(* CODESYS project Controls.export

Project tree, tasks and I/O mapping:
  visualisation Controls
*)

// /Controls
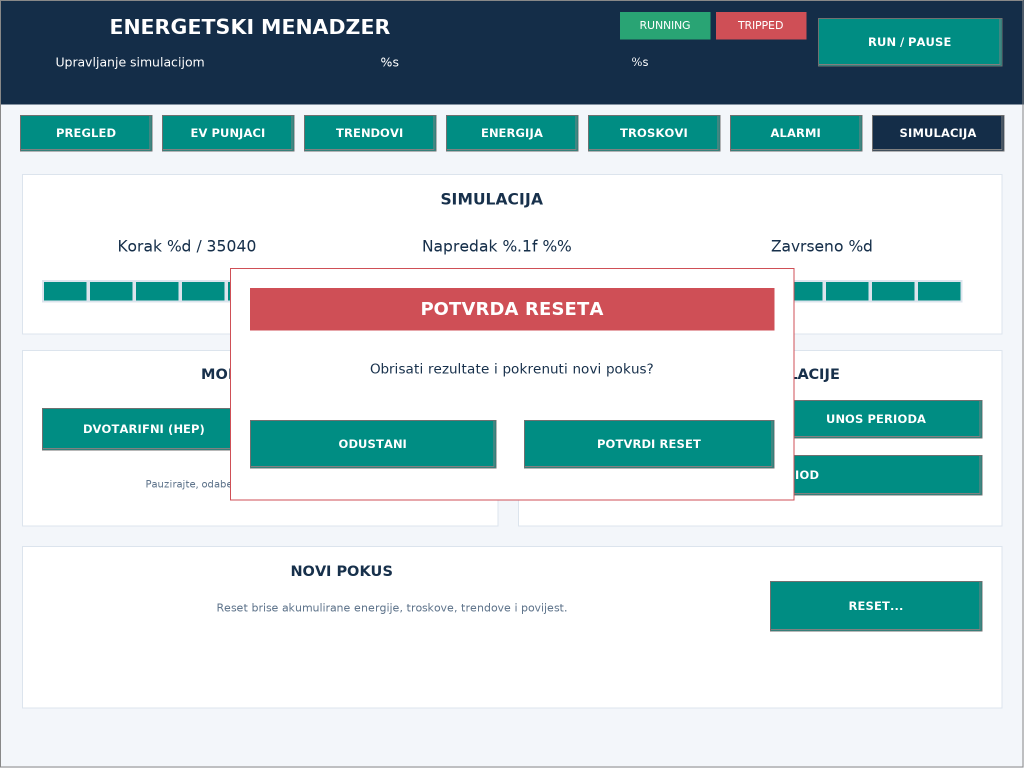
VISUALIZATION Controls  // 1024x768
    Rectangle (0,0 1024x768)
    Rectangle (0,0 1024x104)
    Rectangle (20,10 460x34), "ENERGETSKI MENADZER"
    Rectangle (20,48 220x28), "Upravljanje simulacijom"
    Rectangle (260,49 260x26), "%s", text variable: Team_HMI.sDateTime
    Rectangle (530,49 220x26), "%s", text variable: Team_HMI.sPriceMode
    Button (818,18 184x48), "RUN / PAUSE"
        toggle SimCtrl.run
    Rectangle (620,12 90x27), "PAUSED", invisible if: SimCtrl.run
    Rectangle (620,12 90x27), "RUNNING", invisible if: NOT SimCtrl.run
    Rectangle (716,12 90x27), "TRIPPED", invisible if: NOT SimCtrl.tripped
    Button (20,115 132x36), "PREGLED"
        OnMouseClick:  Assign=Overview, Type=Assignment
    Button (162,115 132x36), "EV PUNJACI"
        OnMouseClick:  Assign=EVs, Type=Assignment
    Button (304,115 132x36), "TRENDOVI"
        OnMouseClick:  Assign=Trends, Type=Assignment
    Button (446,115 132x36), "ENERGIJA"
        OnMouseClick:  Assign=Energy, Type=Assignment
    Button (588,115 132x36), "TROSKOVI"
        OnMouseClick:  Assign=Costs, Type=Assignment
    Button (730,115 132x36), "ALARMI"
        OnMouseClick:  Assign=Alarms, Type=Assignment
    Button (872,115 132x36), "SIMULACIJA"
        OnMouseClick:  Assign=Controls, Type=Assignment
    Rectangle (22,174 980x160)
    Rectangle (42,185 900x28), "SIMULACIJA"
    Rectangle (42,229 290x34), "Korak %d / 35040", text variable: SimCtrl.k
    Rectangle (352,229 290x34), "Napredak %.1f %%", text variable: Team_HMI.rProgressPct
    Rectangle (662,229 320x34), "Zavrseno %d", text variable: BOOL_TO_INT(SimCtrl.finished)
    Rectangle (42,280 920x22)
    Rectangle (44,282 42x18), invisible if: (Team_HMI.rProgressPct) < 5.000
    Rectangle (90,282 42x18), invisible if: (Team_HMI.rProgressPct) < 10.000
    Rectangle (136,282 42x18), invisible if: (Team_HMI.rProgressPct) < 15.000
    Rectangle (182,282 42x18), invisible if: (Team_HMI.rProgressPct) < 20.000
    Rectangle (228,282 42x18), invisible if: (Team_HMI.rProgressPct) < 25.000
    Rectangle (274,282 42x18), invisible if: (Team_HMI.rProgressPct) < 30.000
    Rectangle (320,282 42x18), invisible if: (Team_HMI.rProgressPct) < 35.000
    Rectangle (366,282 42x18), invisible if: (Team_HMI.rProgressPct) < 40.000
    Rectangle (412,282 42x18), invisible if: (Team_HMI.rProgressPct) < 45.000
    Rectangle (458,282 42x18), invisible if: (Team_HMI.rProgressPct) < 50.000
    Rectangle (504,282 42x18), invisible if: (Team_HMI.rProgressPct) < 55.000
    Rectangle (550,282 42x18), invisible if: (Team_HMI.rProgressPct) < 60.000
    Rectangle (596,282 42x18), invisible if: (Team_HMI.rProgressPct) < 65.000
    Rectangle (642,282 42x18), invisible if: (Team_HMI.rProgressPct) < 70.000
    Rectangle (688,282 42x18), invisible if: (Team_HMI.rProgressPct) < 75.000
    Rectangle (734,282 42x18), invisible if: (Team_HMI.rProgressPct) < 80.000
    Rectangle (780,282 42x18), invisible if: (Team_HMI.rProgressPct) < 85.000
    Rectangle (826,282 42x18), invisible if: (Team_HMI.rProgressPct) < 90.000
    Rectangle (872,282 42x18), invisible if: (Team_HMI.rProgressPct) < 95.000
    Rectangle (918,282 42x18), invisible if: (Team_HMI.rProgressPct) < 100.000
    Rectangle (22,350 476x176)
    Rectangle (42,360 436x28), "MODEL CIJENA"
    Button (42,408 204x42), "DVOTARIFNI (HEP)"
        OnMouseClick: execute { IF NOT SimCtrl.run THEN SimCtrl.price_mode := 0; END_IF; }
    Button (262,408 216x42), "DAN UNAPRIJED"
        OnMouseClick: execute { IF NOT SimCtrl.run THEN SimCtrl.price_mode := 1; END_IF; }
    Rectangle (42,470 436x28), "Pauzirajte, odaberite model, zatim resetirajte."
    Rectangle (518,350 484x176)
    Rectangle (538,360 444x28), "BRZINA SIMULACIJE"
    Rectangle (538,400 216x38), "Period: %u ms", text variable: SimCtrl.cycle_time_ms
    Button (770,400 212x38), "UNOS PERIODA"
        OnMouseClick: write SimCtrl.cycle_time_ms via Default, min 10, max 60000, title 'UNOS PERIODA'
    Button (538,455 444x40), "PRIMIJENI PERIOD"
        tap SimCtrl.change_cycle
    Rectangle (22,546 980x162)
    Rectangle (42,557 600x28), "NOVI POKUS"
    Rectangle (42,594 700x28), "Reset brise akumulirane energije, troskove, trendove i povijest."
    Button (770,581 212x50), "RESET..."
        OnMouseClick: execute { Team_Visu.xResetArmed := TRUE; }
    Rectangle (230,268 564x232), invisible if: NOT Team_Visu.xResetArmed
    Rectangle (250,288 524x42), "POTVRDA RESETA", invisible if: NOT Team_Visu.xResetArmed
    Rectangle (250,346 524x46), "Obrisati rezultate i pokrenuti novi pokus?", invisible if: NOT Team_Visu.xResetArmed
    Button (250,420 246x48), "ODUSTANI", invisible if: NOT Team_Visu.xResetArmed
        OnMouseClick: execute { Team_Visu.xResetArmed := FALSE; }
    Button (524,420 250x48), "POTVRDI RESET", invisible if: NOT Team_Visu.xResetArmed
        OnMouseClick: execute { SimCtrl.run := FALSE; SimCtrl.reset := TRUE; Team_Visu.xResetArmed := FALSE; }
END_VISUALIZATION
